(*
SPDX-FileCopyrightText: c 2026 Oleksandr Tiutyk <trofimich@gmail.com>
SPDX-License-Identifier: MIT
License: https://opensource.org/license/mit
*)

(*!
<summary>Checks output writes and acknowledgements of both transitions.</summary>
<description>
Uses a live case-owned automation parent and fresh local device fixtures on every run.
The scenario reads and writes ordinary simulated storage within one task cycle.
</description>
*)

{attribute 'no_assign'}
{attribute 'no_explicit_call' := 'do not call this function block directly'}
FUNCTION_BLOCK DigitalOutputNormallyOpenTest EXTENDS TOF_Testing.SingleCycleTest
VAR_STAT
	{attribute 'hide'}
	_ClassName : STRING := __POUNAME();
END_VAR
VAR
	//! <summary>Live parent borrowed by the method-local simulated device.</summary>
	_AutomationRoot : MockAutomationController(name := "DevicesIORoot");
END_VAR

(*!
<summary>Checks output writes and acknowledgements of both transitions.</summary>
*)
METHOD PROTECTED ExecuteTest
VAR
	output : TOF_Devices_IO.DigitalOutput(name := "DO_NO", parent := _AutomationRoot);
	rawOutput : BOOL;
END_VAR
output.Initialize();
output.BindToIO(rawValue := rawOutput);

output.Value := TRUE;
Assert.ThatBool(
	actual := output.Changed,
	message := "Changed must be TRUE before processing a new value"
).IsTrue();
output.ProcessOutput();
Assert.ThatBool(
	actual := rawOutput,
	message := "rawOutput should be TRUE"
).IsTrue();
Assert.ThatBool(
	actual := output.Changed,
	message := "Processing acknowledges the current value"
).IsFalse();

output.Value := FALSE;
Assert.ThatBool(
	actual := output.Changed,
	message := "The reverse transition must also be pending"
).IsTrue();
output.ProcessOutput();
Assert.ThatBool(
	actual := output.Changed,
	message := "Processing acknowledges the reverse transition"
).IsFalse();
Assert.ThatBool(
	actual := rawOutput,
	message := "rawOutput should be FALSE"
).IsFalse();
END_METHOD

//! <summary>Borrows the concrete class name. Callers must not modify it.</summary>
{attribute 'monitoring' := 'call'}
PROPERTY ClassName : REFERENCE TO STRING
GET
ClassName REF= _ClassName;
END_GET
END_PROPERTY

//! <summary>Borrows the compiler-initialized namespace name. Callers must not modify it.</summary>
{attribute 'monitoring' := 'call'}
PROPERTY NamespaceName : REFERENCE TO STRING
GET
NamespaceName REF= CurrentNamespace.Name;
END_GET
END_PROPERTY

//! <summary>Reports the concrete instance size in bytes.</summary>
{attribute 'monitoring' := 'call'}
PROPERTY SelfSize : ULINT
GET
SelfSize := XSIZEOF(THIS^);
END_GET
END_PROPERTY

END_FUNCTION_BLOCK

(* stored: Version 1.1.0.1
   POU DigitalOutputNormallyOpenTest: Id {22ad81c1-a9ec-4dce-adfa-07da415105ff}, SpecialFunc None
   Method ExecuteTest: Id {d648d6d3-461f-4e8d-a23f-6961d3f8d03a}
   Property ClassName: Id {2a000457-0ff3-45d8-b78b-8f9c6e71148a}
   Get Get: Id {1fedda93-503e-44ee-82a3-d4585134bdc5}
   Property NamespaceName: Id {6ccb5268-5dc6-41b1-a549-cdd84c2f0377}
   Get Get: Id {396cbee8-9b70-45b6-9b44-201e8c768fc5}
   Property SelfSize: Id {db342b77-3b46-4aa7-848c-40544fd0fc55}
   Get Get: Id {027ed52a-4ba8-4185-9d20-6c8815ba666e} *)
